Fanuc KAREL source: KA00161.KL

PROGRAM KA00161
%NOLOCKGROUP
VAR
  SRC: ARRAY[4] OF REAL
  DST: ARRAY[4] OF XYZWPR
BEGIN
  DST = SRC
END KA00161
